FUNCTION_BLOCK CapDistributionCAT (* CAT Function Block Type *)
  (* Standard: 61499-2 *)
  (* Version 0.0, 7/10/2026, template *)
  PACKAGE Main;
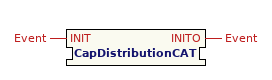
  EVENT_INPUT
    INIT; (* Initialization Request *)
  END_EVENT
  EVENT_OUTPUT
    INITO; (* Initialization Confirm *)
  END_EVENT
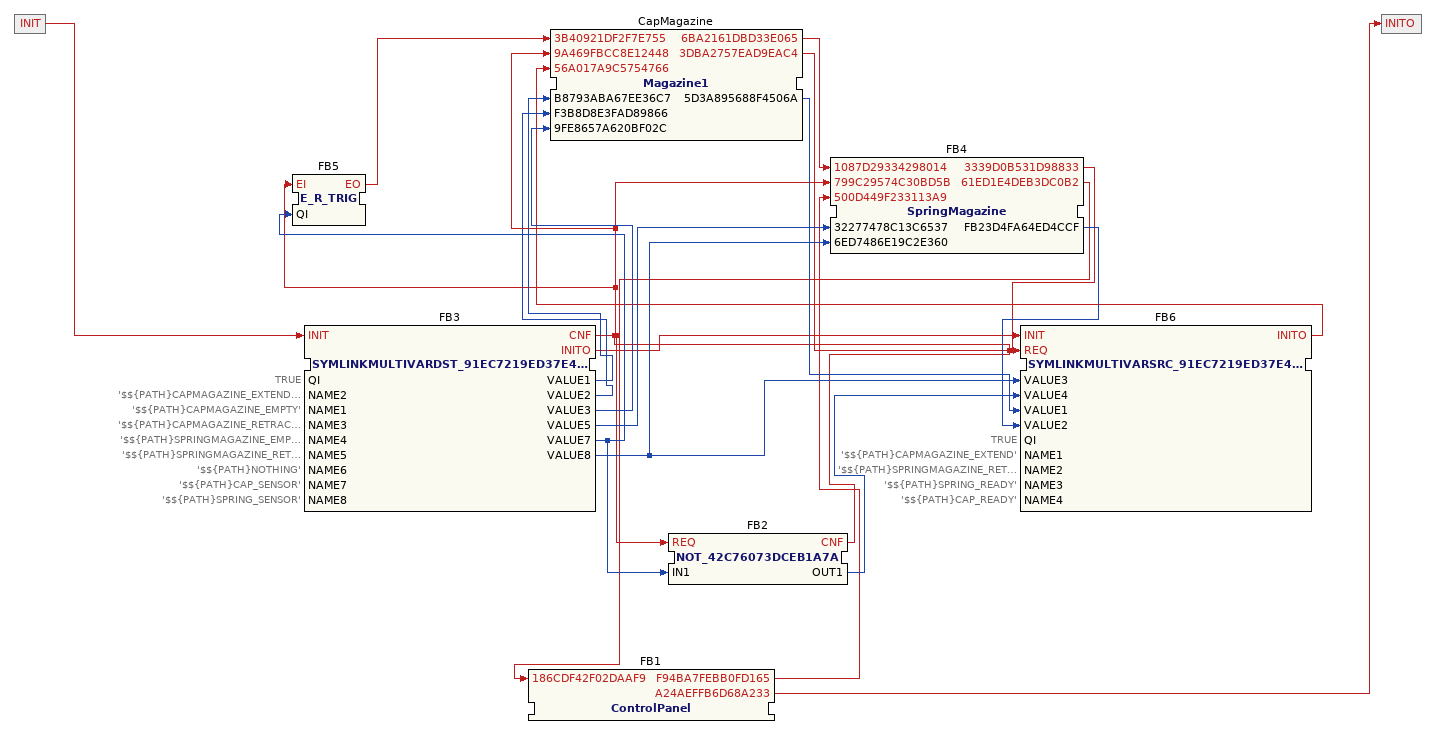
  FBS
    FB1 : ControlPanel;
    FB2 : NOT_42C76073DCEB1A7A; {SET_ATTRIBUTE(Configuration.GenericFBType.InterfaceParams, Runtime.Standard#CNT:=1;OUT${CNT$}:BOOL)}
    CapMagazine : Magazine1;
    FB4 : SpringMagazine;
    FB5 : E_R_TRIG;
    FB6 : SYMLINKMULTIVARSRC_91EC7219ED37E472(QI := TRUE, NAME1 := '$${PATH}CAPMAGAZINE_EXTEND', NAME2 := '$${PATH}SPRINGMAGAZINE_RETRACT', NAME3 := '$${PATH}SPRING_READY', NAME4 := '$${PATH}CAP_READY'); {SET_ATTRIBUTE(Configuration.GenericFBType.InterfaceParams, Runtime.System#I:=8;VALUE${I$}:BOOL,BOOL,BOOL,BOOL,BOOL,BOOL,BOOL,BOOL)}
    FB3 : SYMLINKMULTIVARDST_91EC7219ED37E472(QI := TRUE, NAME2 := '$${PATH}CAPMAGAZINE_EXTENDED', NAME1 := '$${PATH}CAPMAGAZINE_EMPTY', NAME3 := '$${PATH}CAPMAGAZINE_RETRACTED', NAME4 := '$${PATH}SPRINGMAGAZINE_EMPTY', NAME5 := '$${PATH}SPRINGMAGAZINE_RETRACTED', NAME6 := '$${PATH}NOTHING', NAME7 := '$${PATH}CAP_SENSOR', NAME8 := '$${PATH}SPRING_SENSOR'); {SET_ATTRIBUTE(Configuration.GenericFBType.InterfaceParams, Runtime.System#I:=8;VALUE${I$}:BOOL,BOOL,BOOL,BOOL,BOOL,BOOL,BOOL,BOOL)}
  END_FBS
  EVENT_CONNECTIONS
    FB5.EO TO CapMagazine.3B40921DF2F7E755;
    CapMagazine.6BA2161DBD33E065 TO FB4.1087D29334298014;
    INIT TO FB3.INIT;
    FB3.CNF TO FB5.EI;
    FB3.CNF TO CapMagazine.9A469FBCC8E12448;
    FB3.CNF TO FB4.799C29574C30BD5B;
    FB3.CNF TO FB2.REQ;
    FB3.INITO TO FB6.INIT;
    CapMagazine.3DBA2757EAD9EAC4 TO FB6.REQ;
    FB4.3339D0B531D98833 TO FB6.REQ;
    FB2.CNF TO FB6.REQ;
    FB3.CNF TO FB6.REQ;
    FB6.INITO TO CapMagazine.56A017A9C5754766;
    FB4.61ED1E4DEB3DC0B2 TO FB1.186CDF42F02DAAF9;
    FB1.F94BA7FEBB0FD165 TO FB4.500D449F233113A9;
    FB1.A24AEFFB6D68A233 TO INITO;
  END_CONNECTIONS
  DATA_CONNECTIONS
    FB3.VALUE1 TO CapMagazine.B8793ABA67EE36C7;
    FB3.VALUE2 TO CapMagazine.F3B8D8E3FAD89866;
    FB3.VALUE3 TO CapMagazine.9FE8657A620BF02C;
    FB3.VALUE5 TO FB4.32277478C13C6537;
    FB3.VALUE7 TO FB2.IN1;
    FB3.VALUE7 TO FB5.QI;
    FB3.VALUE8 TO FB6.VALUE3;
    FB3.VALUE8 TO FB4.6ED7486E19C2E360;
    FB2.OUT1 TO FB6.VALUE4;
    CapMagazine.5D3A895688F4506A TO FB6.VALUE1;
    FB4.FB23D4FA64ED4CCF TO FB6.VALUE2;
  END_CONNECTIONS
END_FUNCTION_BLOCK
